FUNCTION_BLOCK FB_Hysteresis_REAL
VAR_INPUT
	fIn		: REAL; // in case of iDigitsAfterDot=2 max value 327.67 * 100 >> INTEGER Value limitation
	fHigh	: REAL;
	fLow	: REAL;
	iDigitsAfterDot: INT:=1; //min 0 , max 3

END_VAR
VAR_OUTPUT
	bOut	: BOOL;
END_VAR
VAR
	fbHys: HYSTERESIS;
	mult: INT;
	iDigitsAfterDot_Local: INT:=2; //min 0 , max 3


END_VAR

IF iDigitsAfterDot < 0 THEN;
	iDigitsAfterDot_Local:=0;
ELSIF iDigitsAfterDot > 3 THEN;
	iDigitsAfterDot_Local:=3;
ELSE;
	iDigitsAfterDot_Local:=iDigitsAfterDot;
END_IF
 

CASE iDigitsAfterDot_Local OF
	0:mult:=1;
	1:mult:=10;
	2:mult:=100;
	3:mult:=1000;
END_CASE

fbHys.HIGH:=REAL_TO_INT(fHigh*mult);
fbHys.LOW:=REAL_TO_INT(fLow*mult);
fbHys.IN:=REAL_TO_INT(fIn*mult);

fbHys(OUT=>bOut);

END_FUNCTION_BLOCK

(* stored: Version 1.1.0.1, ProductVersion 3.1.4024.12
   POU FB_Hysteresis_REAL: Id {db4e44f4-3d76-460f-ab24-9469a97bf7d8}, SpecialFunc None *)
